(* IEC 61131-3 sources: CannyIECUnitTest/st/device/plc_logic/application/testcase_isignbit, 1 file *)

(* ---- execute-Execute.st ---- *)
(* --- Interface --- *)
METHOD PROTECTED Execute : BOOL
VAR_OUTPUT
	iErrorCode : INT;
END_VAR
VAR
	xAssert : BOOL;
END_VAR

(* --- Implementation --- *)
xAssert := TM.Assert_Bool_IsFalse(context := THIS^, actualValue := CANNY.ISIGNBIT(0), wsErrorMsg := "");
xAssert := TM.Assert_Bool_IsTrue(context := THIS^, actualValue := CANNY.ISIGNBIT(-1), wsErrorMsg := "");
xAssert := TM.Assert_Bool_IsFalse(context := THIS^, actualValue := CANNY.ISIGNBIT(1), wsErrorMsg := "");
Execute := TRUE;
